Fanuc KAREL source: kx00033.compact.KL

PROGRAM KX00033
%STACKSIZE=65535
%PRIORITY=65535
%UNINITVARS
%NOLOCKGROUP
VAR
I : INTEGER
J : INTEGER
B : BOOLEAN
F : FILE
S : STRING[80]
P : XYZWPR
BEGIN
I=1
END KX00033
